// TIA Portal V21 export
// export: Created 2026-11-10T19:13:03.1555193Z, ExportSetting WithDefaults, DisplayName Totally Integrated Automation Portal, DisplayVersion V21 Update 3, DisplayName STEP 7 Professional, DisplayVersion V21 Update 3, DisplayName STEP 7 Safety, DisplayVersion V21, DisplayName Tech WebApplication, DisplayVersion V21, DisplayName WinCC Basic/Comfort/Advanced, DisplayVersion V21 Update 3, DisplayName WinCC Unified, DisplayVersion V21 Update 3
FUNCTION "FC_TsendB" : Void   // FC4, SCL
{ S7_Optimized_Access := 'TRUE' }
VERSION : 0.1
// stored: AutoNumber true, IsIECCheckEnabled false, SetENOAutomatically false, UDAEnableTagReadback false
BEGIN
   "DB_TSEND".TSEND(REQ := FALSE, ID := W#16#1, LEN := 0, DATA := "DB_Buf".buf); "DB_TRCV".TRCV(EN_R := FALSE, ID := W#16#1, LEN := 0, DATA := "DB_Buf".buf);
END_FUNCTION
